(* IEC 61131-3 sources: SRCI_CLIENT_PLC/RobotLibrary/Library/Structures/AxesGroup/State/DataChanged, 1 file *)

(* ---- AxesGroupStateDataChanged.st ---- *)
{attribute 'pack_mode' := '1'}
// -------------------------------------------------------------------------
//  SRCI Robot Library
// -------------------------------------------------------------------------
//
//  Object:      AxesGroupStateDataChanged
//  Author:      Thorsten Brach
//  Date:        2024-06-01
//
//  Description:
//
//
//  Copyright:
//    (C) 2024 Thorsten Brach. All rights reserved
//             Licensed under the MIT License.
//
//  Disclaimer:
//    This project is provided without any guarantee and can be used for
//    private and commercial purposes. Any use is at the user’s
//    own risk and responsibility.
//
// -------------------------------------------------------------------------
TYPE AxesGroupStateDataChanged :
STRUCT
  /// indicates that tool data has changed
  Tool              : ARRAY[0..RobotLibraryParameter.TOOL_MAX       -1] OF BOOL;
  /// indicates that frame data has changed
  Frame             : ARRAY[0..RobotLibraryParameter.FRAME_MAX      -1] OF BOOL;
  /// indicates that load data has changed
  Load              : ARRAY[0..RobotLibraryParameter.LOAD_MAX       -1] OF BOOL;
  /// indicates that work area has changed
  WorkArea          : ARRAY[0..RobotLibraryParameter.WORK_AREAS_MAX -1] OF BOOL;
  /// indicates that default dynamic has changed
  DefaultDynamics   : BOOL;
  /// indicates that reference dynamic has changed
  ReferenceDynamics : BOOL;
  /// indicates that software limits has changed
  SwLimits          : BOOL;
END_STRUCT
END_TYPE
